VAR_GLOBAL
    enabled : ARRAY[1..3] OF BOOL := [TRUE, TRUE, TRUE];
    sensor : ARRAY[1..3] OF BOOL;
    blocked : ARRAY[1..3] OF BOOL;
    running : ARRAY[1..3] OF BOOL;
    actualSpeed : ARRAY[1..3] OF REAL;
    productCount : ARRAY[1..3] OF DINT;
    alarm : ARRAY[1..3] OF STRING(80);
END_VAR

(* stored: Version 1.1.0.1, ProductVersion 3.1 *)
